// FC_INT_TO_TIME: INT转TIME (占位版本)
// 描述: 在LSP环境中返回T#0ms, 避免类型转换错误

FUNCTION FC_INT_TO_TIME : TIME
VAR_INPUT
    IntValue : INT;
END_VAR

BEGIN
    // [多平台占位] LSP环境返回T#0ms
    FC_INT_TO_TIME := T#0ms;

END_FUNCTION
